(* PLC project Vn_sr_call, Beckhoff Automation GmbH TwinCAT PLC Control 3.5.13.21 *)
(* stored: creationDateTime 1970-01-01T00:00:00 *)

PROGRAM Vn_sr_call

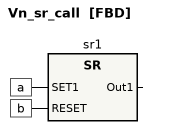
(* FBD diagram, written out as Structured Text *)
sr1(SET1 := a, RESET := b);
END_PROGRAM
